TYPE "ST_AirPressureHal"
VERSION : 0.1
   STRUCT
      LowPressure : Bool;
      OperatingPressure : Bool;
      Quality : Bool := TRUE;
   END_STRUCT;

END_TYPE

